(* IEC 61131-3 sources: rusty/tests/integration/data/linking, 7 files *)

(* ---- init.st ---- *)
TYPE myStruct : STRUCT
    a : INT := 5;
    b : DINT := 6;
END_STRUCT
END_TYPE

(* ---- consts.st ---- *)
VAR_GLOBAL CONSTANT
    myValue : BOOL := TRUE;
END_VAR

FUNCTION main : DINT
END_FUNCTION

(* ---- file1.st ---- *)
{external}
FUNCTION func2 : DINT
END_FUNCTION

FUNCTION func1 : DINT
    func2();
END_FUNCTION

(* ---- file2.st ---- *)
{external}
FUNCTION func1 : DINT
END_FUNCTION

FUNCTION func2 : DINT
    func1();
END_FUNCTION

(* ---- relative.st ---- *)
FUNCTION relative : DINT
END_FUNCTION

(* ---- init2.st ---- *)
FUNCTION_BLOCK myFB
    VAR
        myS : myStruct := (a := 2);
    END_VAR
END_FUNCTION_BLOCK

(* ---- init3.st ---- *)
FUNCTION_BLOCK myFb2
    VAR
        fb : myFb;
    END_VAR
END_FUNCTION_BLOCK
